// TIA Portal V21 program export: 1 tag tables, 0 data types, 0 data blocks, 4 code blocks (in call order from the OBs), 1 instance data blocks

VAR_GLOBAL   // PLC tag table "Default tag table"
END_VAR

ORGANIZATION_BLOCK "Main"   // OB1, SCL, ProgramCycle
{ S7_Optimized_Access := 'TRUE' }
VERSION : 0.1
// stored: AutoNumber true, IsIECCheckEnabled false, SetENOAutomatically false
   VAR_INPUT
      Initial_Call : Bool;   // Initial call of this OB
      Remanence : Bool;   // =True, if remanent data are available
   END_VAR
BEGIN
      "TiaMcp_EnableGate_DB"(Enable := TRUE);
END_ORGANIZATION_BLOCK

FUNCTION_BLOCK "TiaMcp_EnableGate"   // FB1, SCL
{ S7_Optimized_Access := 'TRUE' }
VERSION : 0.1
// stored: AutoNumber true, IsIECCheckEnabled false, IsRetainMemResEnabled false, MemoryReserve 100, SetENOAutomatically false, UDAEnableTagReadback false
   VAR_INPUT
      Enable : Bool;
   END_VAR
   VAR_OUTPUT
      Active : Bool;
   END_VAR
BEGIN
      #Active := "TiaMcp_IsEnabled"(Enable := #Enable);
END_FUNCTION_BLOCK

FUNCTION "TiaMcp_IsEnabled" : Bool   // FC1, SCL
{ S7_Optimized_Access := 'TRUE' }
VERSION : 0.1
// stored: AutoNumber true, IsIECCheckEnabled false, SetENOAutomatically false, UDAEnableTagReadback false
   VAR_INPUT
      Enable : Bool;
   END_VAR
BEGIN
      #TiaMcp_IsEnabled := #Enable;
END_FUNCTION

BLOCK "Force table"   // PlcForceTable
BEGIN
END_BLOCK

DATA_BLOCK "TiaMcp_EnableGate_DB"   // DB1
VERSION : 0.1
// stored: AutoNumber true, DBAccessibleFromOPCUA true, DBAccessibleFromWebserver true, InstanceOfName TiaMcp_EnableGate, InstanceOfType FB
"TiaMcp_EnableGate"
BEGIN
END_DATA_BLOCK
